TYPE ST_HeatExchanger :
STRUCT
	//request
	bManual	:	BOOL	;//System in automatic
	bRun	:	BOOL	;
	nTemp	:	INT		;
	//feedback
	nTemp_fdbk	:	INT	;
	
	//Output signal scaling
	cntrlVal_Min		: REAL:=0;
	cntrlVal_Max		: REAL:=100;
	
	outVal_Min		: REAL:=0;
	outVal_Max		: REAL:=32767;
	outOffset		: REAL:=0;
	fManualControl	: LREAL:=100;

END_STRUCT
END_TYPE

(* stored: Version 1.1.0.1, ProductVersion 3.1.4024.13
   DUT ST_HeatExchanger: Id {fdaef3e3-531e-423e-9e26-9ca260edffe0} *)
